(* IEC 61131-3 sources: axsharp/src/ix.connectors/tests/ax-test-project/src/issues, 1 file *)

(* ---- GH-PKTu-ix_56.st ---- *)
// https://github.com/ix-ax/ix/issues/56
NAMESPACE GH.PKTu.ix_56

    CLASS ComplexMember
        VAR PUBLIC
            Counter : INT;
        END_VAR

    END_CLASS

    CLASS Base
        VAR PUBLIC
            baseMember : STRING;
            baseComplexMember : ComplexMember;
            BaseDavid : DavidBase;
        END_VAR
    END_CLASS

    CLASS FirstInheritance EXTENDS Base
        VAR PUBLIC
            FirstInheritanceMember : STRING;
            FirstInheritanceComplexMember : ComplexMember;
            FirstDavid : DavidBase;
        END_VAR
    END_CLASS

    CLASS SecondInheritance EXTENDS FirstInheritance
        VAR PUBLIC
            SecondInheritanceMember : STRING;
            SecondInheritanceComplexMember : ComplexMember;
            SecodnDavid : DavidBase;
        END_VAR
    END_CLASS

    CLASS PedroBase
        VAR PUBLIC
            p : STRING;
        END_VAR
    END_CLASS

    CLASS DavidBase EXTENDS PedroBase
        VAR PUBLIC
            d : STRING;
        END_VAR
    END_CLASS
END_NAMESPACE
